// TIA Portal V17 export
// export: Created 2025-08-05T06:59:04.9381121Z, ExportSetting WithDefaults, DisplayName Totally Integrated Automation Portal, DisplayVersion V17 Update 5, DisplayName TIA Portal Openness, DisplayVersion V17 Update 5, DisplayName TIA Portal Version Control Interface, DisplayVersion V17, DisplayName SINAMICS Startdrive Advanced, DisplayVersion V17, DisplayName SINAMICS Startdrive G130, G150, S120, S150, SINAMICS MV, S210, DisplayVersion V17, DisplayName SINAMICS Startdrive G110M, G120, G120C, G120D, G120P, G115D, DisplayVersion V17, DisplayName STEP 7 Professional, DisplayVersion V17 Update 5, DisplayName STEP 7 Safety, DisplayVersion V17, DisplayName WinCC Advanced, DisplayVersion V17 Update 5
FUNCTION_BLOCK "FB_CentreStand_Fix_Seq_7"   // FB1, LAD
VERSION : 0.1
// stored: AutoNumber true, IsIECCheckEnabled false, UDAEnableTagReadback false
   VAR_INPUT
      iAutoRunning : Bool;
      iFixClamp : Bool;
      iFixEmpty : Bool;
      iFixTrayPresent : Bool;
      iFixUnclamp : Bool;
      iR1DropOver : Bool;
      iR1PickOver : Bool;
      iR2OperationOver : Bool;
      iR2ServiceActivated : Bool;
      iR2ServiceCompleted : Bool;
      iReset_fault : Bool;
      iRobotOutofZone : Bool;
      iSstMode : Bool;
      iSstPB : Bool;
   END_VAR
   VAR_OUTPUT
      qFixClamp : Bool;
      qFixUnclamp : Bool;
      qR1ReadytoDropTray : Bool;
      qR1ReadytoPickTray : Bool;
      qR2OperationStart : Bool;
   END_VAR
   VAR_IN_OUT
      iqR2ServiceActive : Bool;
      iqR2ServiceCompleted : Bool;
   END_VAR
   VAR DB_SPECIFIC
      StateNo : Int;
      s138_WaitBothRbtOutAl : Bool;
      s138_WaitBothRbtOutAl_T1 : Bool;
      s138_WaitBothRbtOutAl_T2 : Bool;
      s139_FixEmpty : Bool;
      s139_FixEmpty_T1 : Bool;
      s140_FixTrayPrsntRec : Bool;
      s140_FixTrayPrsntRec_T1 : Bool;
      s140_FixTrayPrsntRec_T2 : Bool;
      s141_FixUnclampCmd : Bool;
      s141_FixUnclampCmd_T1 : Bool;
      s142_TrayRdyDropFix : Bool;
      s142_TrayRdyDropFix_T1 : Bool;
      s143_RbtDropFixChkTr : Bool;
      s143_RbtDropFixChkTr_T1 : Bool;
      s144_RbtOutAreaDrop : Bool;
      s144_RbtOutAreaDrop_T1 : Bool;
      s145_FixClamp : Bool;
      s145_FixClamp_T1 : Bool;
      s146_Rbt2AlloyOpOver : Bool;
      s146_Rbt2AlloyOpOver_T1 : Bool;
      s147_FixUnclmpCmdOvr : Bool;
      s147_FixUnclmpCmdOvr_T1 : Bool;
      s148_RdyPickTrayWait : Bool;
      s148_RdyPickTrayWait_T1 : Bool;
      s149_RbtPickTrayChkEm : Bool;
      s149_RbtPickTrayChkEm_T1 : Bool;
      s191_WaitRbt2OutArea : Bool;
      s191_WaitRbt2OutArea_T1 : Bool;
      sSst : Bool;
      sSstPulse : Bool;
      sSstRise : Bool;
      sStWtResetRel : Bool;
      sStWtResetRel_T1 : Bool;
   END_VAR
   VAR_TEMP
      tOne : Bool;
   END_VAR
   VAR_TEMP   // added for the SCL form of the ladder/FBD networks
      _w1 : Bool;
   END_VAR
BEGIN

REGION Network 1
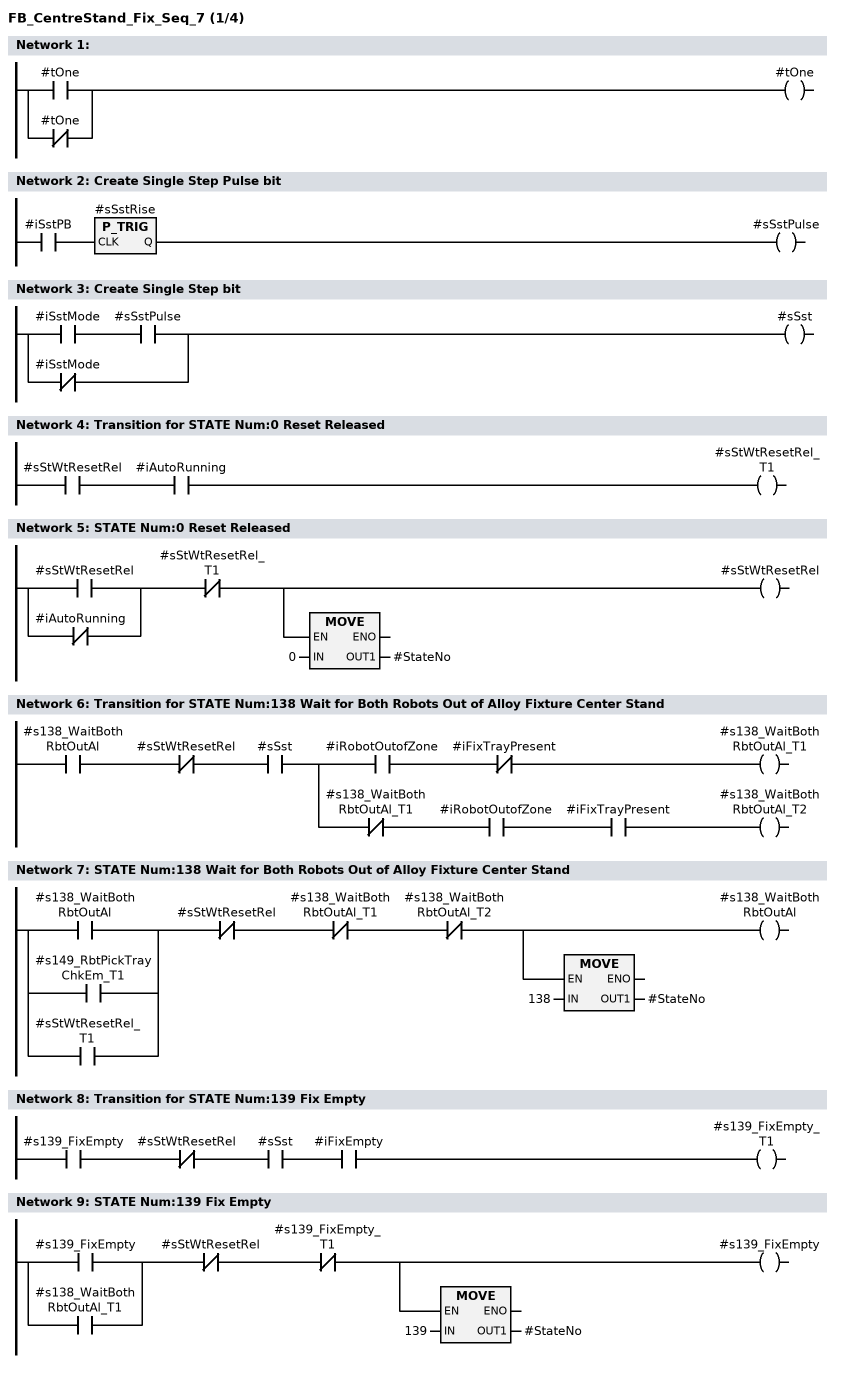
   RUNG wire#powerrail
      Contact( #tOne )
      wire#w1
      Coil( #tOne )
   END_RUNG
   RUNG wire#powerrail
      I_Contact( #tOne )
   END_RUNG wire#w1
   // the same network as SCL:
   #tOne := #tOne OR NOT #tOne;
END_REGION

REGION Network 2: Create Single Step Pulse bit
   RUNG wire#powerrail
      Contact( #iSstPB )
      P_Trig( #sSstRise )
      Coil( #sSstPulse )
   END_RUNG
   // the same network as SCL:
   #_w1 := #iSstPB AND NOT #sSstRise;   // rising edge
   #sSstRise := #iSstPB;
   #sSstPulse := #_w1;
END_REGION

REGION Network 3: Create Single Step bit
   RUNG wire#powerrail
      Contact( #iSstMode )
      Contact( #sSstPulse )
      wire#w1
      Coil( #sSst )
   END_RUNG
   RUNG wire#powerrail
      I_Contact( #iSstMode )
   END_RUNG wire#w1
   // the same network as SCL:
   #sSst := (#iSstMode AND #sSstPulse) OR NOT #iSstMode;
END_REGION

REGION Network 4: Transition for STATE Num:0 Reset Released
   RUNG wire#powerrail
      Contact( #sStWtResetRel )
      Contact( #iAutoRunning )
      Coil( #sStWtResetRel_T1 )
   END_RUNG
   // the same network as SCL:
   #sStWtResetRel_T1 := #sStWtResetRel AND #iAutoRunning;
END_REGION

REGION Network 5: STATE Num:0 Reset Released
   RUNG wire#powerrail
      Contact( #sStWtResetRel )
      wire#w1
      I_Contact( #sStWtResetRel_T1 )
      wire#w2
      Coil( #sStWtResetRel )
   END_RUNG
   RUNG wire#powerrail
      I_Contact( #iAutoRunning )
   END_RUNG wire#w1
   RUNG wire#w2
      { S7_GenerateENO := "TRUE" } Move(in := 0, out1 => #StateNo)
   END_RUNG
   // the same network as SCL:
   #sStWtResetRel := (#sStWtResetRel OR NOT #iAutoRunning) AND NOT #sStWtResetRel_T1;
   IF #sStWtResetRel THEN #StateNo := 0; END_IF;
END_REGION

REGION Network 6: Transition for STATE Num:138 Wait for Both Robots Out of Alloy Fixture Center Stand
   RUNG wire#powerrail
      Contact( #s138_WaitBothRbtOutAl )
      I_Contact( #sStWtResetRel )
      Contact( #sSst )
      wire#w1
      Contact( #iRobotOutofZone )
      I_Contact( #iFixTrayPresent )
      Coil( #s138_WaitBothRbtOutAl_T1 )
   END_RUNG
   RUNG wire#w1
      I_Contact( #s138_WaitBothRbtOutAl_T1 )
      Contact( #iRobotOutofZone )
      Contact( #iFixTrayPresent )
      Coil( #s138_WaitBothRbtOutAl_T2 )
   END_RUNG
   // the same network as SCL:
   #_w1 := #s138_WaitBothRbtOutAl AND NOT #sStWtResetRel AND #sSst;
   #s138_WaitBothRbtOutAl_T1 := #_w1 AND #iRobotOutofZone AND NOT #iFixTrayPresent;
   #s138_WaitBothRbtOutAl_T2 := #_w1 AND NOT #s138_WaitBothRbtOutAl_T1 AND #iRobotOutofZone AND #iFixTrayPresent;
END_REGION

REGION Network 7: STATE Num:138 Wait for Both Robots Out of Alloy Fixture Center Stand
   RUNG wire#powerrail
      Contact( #s138_WaitBothRbtOutAl )
      wire#w1
      I_Contact( #sStWtResetRel )
      I_Contact( #s138_WaitBothRbtOutAl_T1 )
      I_Contact( #s138_WaitBothRbtOutAl_T2 )
      wire#w2
      Coil( #s138_WaitBothRbtOutAl )
   END_RUNG
   RUNG wire#powerrail
      Contact( #s149_RbtPickTrayChkEm_T1 )
   END_RUNG wire#w1
   RUNG wire#powerrail
      Contact( #sStWtResetRel_T1 )
   END_RUNG wire#w1
   RUNG wire#w2
      { S7_GenerateENO := "TRUE" } Move(in := 138, out1 => #StateNo)
   END_RUNG
   // the same network as SCL:
   #s138_WaitBothRbtOutAl := (#s138_WaitBothRbtOutAl OR #s149_RbtPickTrayChkEm_T1 OR #sStWtResetRel_T1) AND NOT #sStWtResetRel AND NOT #s138_WaitBothRbtOutAl_T1 AND NOT #s138_WaitBothRbtOutAl_T2;
   IF #s138_WaitBothRbtOutAl THEN #StateNo := 138; END_IF;
END_REGION

REGION Network 8: Transition for STATE Num:139 Fix Empty
   RUNG wire#powerrail
      Contact( #s139_FixEmpty )
      I_Contact( #sStWtResetRel )
      Contact( #sSst )
      Contact( #iFixEmpty )
      Coil( #s139_FixEmpty_T1 )
   END_RUNG
   // the same network as SCL:
   #s139_FixEmpty_T1 := #s139_FixEmpty AND NOT #sStWtResetRel AND #sSst AND #iFixEmpty;
END_REGION

REGION Network 9: STATE Num:139 Fix Empty
   RUNG wire#powerrail
      Contact( #s139_FixEmpty )
      wire#w1
      I_Contact( #sStWtResetRel )
      I_Contact( #s139_FixEmpty_T1 )
      wire#w2
      Coil( #s139_FixEmpty )
   END_RUNG
   RUNG wire#powerrail
      Contact( #s138_WaitBothRbtOutAl_T1 )
   END_RUNG wire#w1
   RUNG wire#w2
      { S7_GenerateENO := "TRUE" } Move(in := 139, out1 => #StateNo)
   END_RUNG
   // the same network as SCL:
   #s139_FixEmpty := (#s139_FixEmpty OR #s138_WaitBothRbtOutAl_T1) AND NOT #sStWtResetRel AND NOT #s139_FixEmpty_T1;
   IF #s139_FixEmpty THEN #StateNo := 139; END_IF;
END_REGION

REGION Network 10: Transition for STATE Num:140 Fix Tray Present_Rec Operation pending
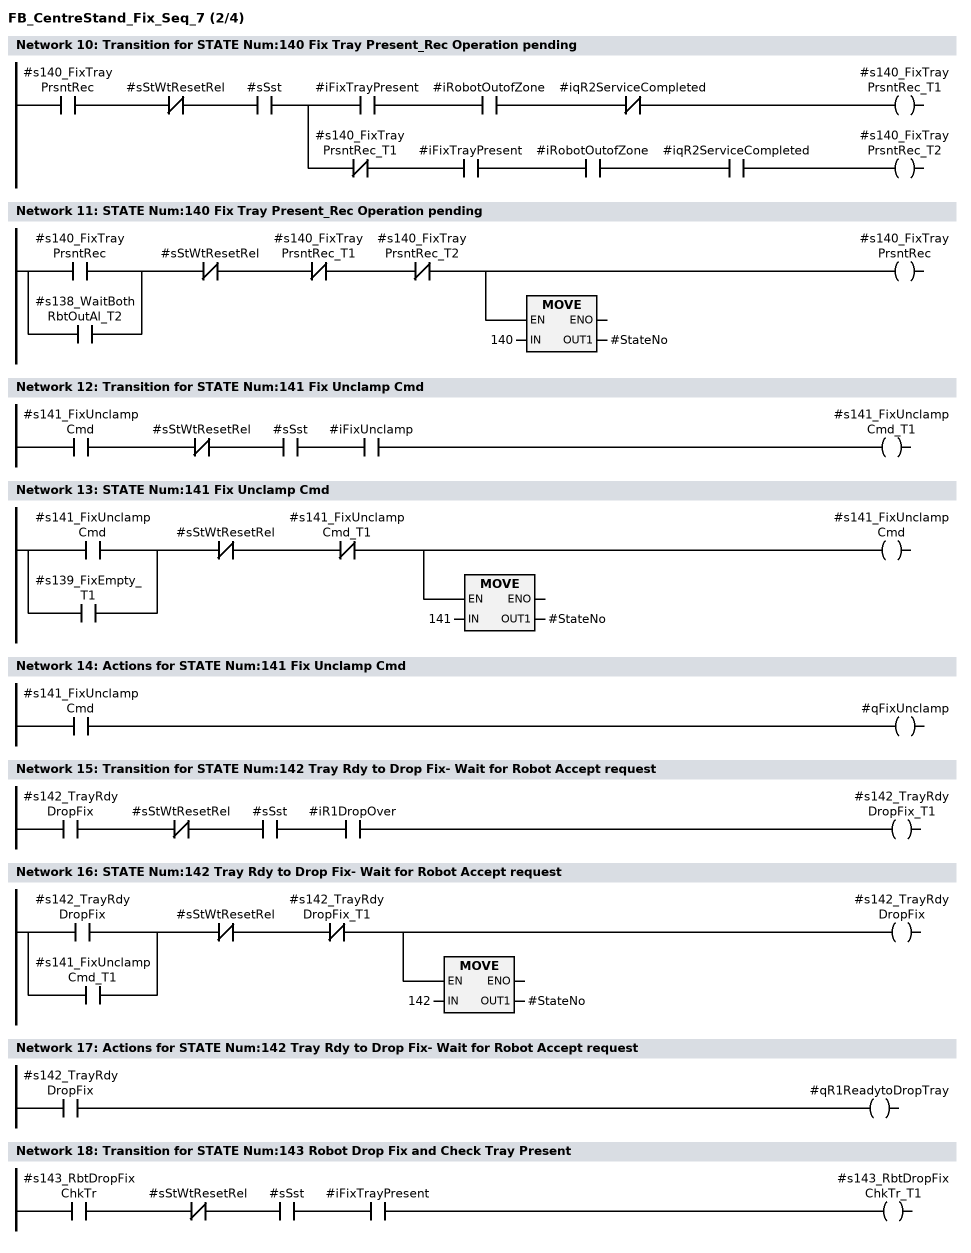
   RUNG wire#powerrail
      Contact( #s140_FixTrayPrsntRec )
      I_Contact( #sStWtResetRel )
      Contact( #sSst )
      wire#w1
      Contact( #iFixTrayPresent )
      Contact( #iRobotOutofZone )
      I_Contact( #iqR2ServiceCompleted )
      Coil( #s140_FixTrayPrsntRec_T1 )
   END_RUNG
   RUNG wire#w1
      I_Contact( #s140_FixTrayPrsntRec_T1 )
      Contact( #iFixTrayPresent )
      Contact( #iRobotOutofZone )
      Contact( #iqR2ServiceCompleted )
      Coil( #s140_FixTrayPrsntRec_T2 )
   END_RUNG
   // the same network as SCL:
   #_w1 := #s140_FixTrayPrsntRec AND NOT #sStWtResetRel AND #sSst;
   #s140_FixTrayPrsntRec_T1 := #_w1 AND #iFixTrayPresent AND #iRobotOutofZone AND NOT #iqR2ServiceCompleted;
   #s140_FixTrayPrsntRec_T2 := #_w1 AND NOT #s140_FixTrayPrsntRec_T1 AND #iFixTrayPresent AND #iRobotOutofZone AND #iqR2ServiceCompleted;
END_REGION

REGION Network 11: STATE Num:140 Fix Tray Present_Rec Operation pending
   RUNG wire#powerrail
      Contact( #s140_FixTrayPrsntRec )
      wire#w1
      I_Contact( #sStWtResetRel )
      I_Contact( #s140_FixTrayPrsntRec_T1 )
      I_Contact( #s140_FixTrayPrsntRec_T2 )
      wire#w2
      Coil( #s140_FixTrayPrsntRec )
   END_RUNG
   RUNG wire#powerrail
      Contact( #s138_WaitBothRbtOutAl_T2 )
   END_RUNG wire#w1
   RUNG wire#w2
      { S7_GenerateENO := "TRUE" } Move(in := 140, out1 => #StateNo)
   END_RUNG
   // the same network as SCL:
   #s140_FixTrayPrsntRec := (#s140_FixTrayPrsntRec OR #s138_WaitBothRbtOutAl_T2) AND NOT #sStWtResetRel AND NOT #s140_FixTrayPrsntRec_T1 AND NOT #s140_FixTrayPrsntRec_T2;
   IF #s140_FixTrayPrsntRec THEN #StateNo := 140; END_IF;
END_REGION

REGION Network 12: Transition for STATE Num:141 Fix Unclamp Cmd
   RUNG wire#powerrail
      Contact( #s141_FixUnclampCmd )
      I_Contact( #sStWtResetRel )
      Contact( #sSst )
      Contact( #iFixUnclamp )
      Coil( #s141_FixUnclampCmd_T1 )
   END_RUNG
   // the same network as SCL:
   #s141_FixUnclampCmd_T1 := #s141_FixUnclampCmd AND NOT #sStWtResetRel AND #sSst AND #iFixUnclamp;
END_REGION

REGION Network 13: STATE Num:141 Fix Unclamp Cmd
   RUNG wire#powerrail
      Contact( #s141_FixUnclampCmd )
      wire#w1
      I_Contact( #sStWtResetRel )
      I_Contact( #s141_FixUnclampCmd_T1 )
      wire#w2
      Coil( #s141_FixUnclampCmd )
   END_RUNG
   RUNG wire#powerrail
      Contact( #s139_FixEmpty_T1 )
   END_RUNG wire#w1
   RUNG wire#w2
      { S7_GenerateENO := "TRUE" } Move(in := 141, out1 => #StateNo)
   END_RUNG
   // the same network as SCL:
   #s141_FixUnclampCmd := (#s141_FixUnclampCmd OR #s139_FixEmpty_T1) AND NOT #sStWtResetRel AND NOT #s141_FixUnclampCmd_T1;
   IF #s141_FixUnclampCmd THEN #StateNo := 141; END_IF;
END_REGION

REGION Network 14: Actions for STATE Num:141 Fix Unclamp Cmd
   RUNG wire#powerrail
      Contact( #s141_FixUnclampCmd )
      Coil( #qFixUnclamp )
   END_RUNG
   // the same network as SCL:
   #qFixUnclamp := #s141_FixUnclampCmd;
END_REGION

REGION Network 15: Transition for STATE Num:142 Tray Rdy to Drop Fix- Wait for Robot Accept request
   RUNG wire#powerrail
      Contact( #s142_TrayRdyDropFix )
      I_Contact( #sStWtResetRel )
      Contact( #sSst )
      Contact( #iR1DropOver )
      Coil( #s142_TrayRdyDropFix_T1 )
   END_RUNG
   // the same network as SCL:
   #s142_TrayRdyDropFix_T1 := #s142_TrayRdyDropFix AND NOT #sStWtResetRel AND #sSst AND #iR1DropOver;
END_REGION

REGION Network 16: STATE Num:142 Tray Rdy to Drop Fix- Wait for Robot Accept request
   RUNG wire#powerrail
      Contact( #s142_TrayRdyDropFix )
      wire#w1
      I_Contact( #sStWtResetRel )
      I_Contact( #s142_TrayRdyDropFix_T1 )
      wire#w2
      Coil( #s142_TrayRdyDropFix )
   END_RUNG
   RUNG wire#powerrail
      Contact( #s141_FixUnclampCmd_T1 )
   END_RUNG wire#w1
   RUNG wire#w2
      { S7_GenerateENO := "TRUE" } Move(in := 142, out1 => #StateNo)
   END_RUNG
   // the same network as SCL:
   #s142_TrayRdyDropFix := (#s142_TrayRdyDropFix OR #s141_FixUnclampCmd_T1) AND NOT #sStWtResetRel AND NOT #s142_TrayRdyDropFix_T1;
   IF #s142_TrayRdyDropFix THEN #StateNo := 142; END_IF;
END_REGION

REGION Network 17: Actions for STATE Num:142 Tray Rdy to Drop Fix- Wait for Robot Accept request
   RUNG wire#powerrail
      Contact( #s142_TrayRdyDropFix )
      Coil( #qR1ReadytoDropTray )
   END_RUNG
   // the same network as SCL:
   #qR1ReadytoDropTray := #s142_TrayRdyDropFix;
END_REGION

REGION Network 18: Transition for STATE Num:143 Robot Drop Fix and Check Tray Present
   RUNG wire#powerrail
      Contact( #s143_RbtDropFixChkTr )
      I_Contact( #sStWtResetRel )
      Contact( #sSst )
      Contact( #iFixTrayPresent )
      Coil( #s143_RbtDropFixChkTr_T1 )
   END_RUNG
   // the same network as SCL:
   #s143_RbtDropFixChkTr_T1 := #s143_RbtDropFixChkTr AND NOT #sStWtResetRel AND #sSst AND #iFixTrayPresent;
END_REGION

REGION Network 19: STATE Num:143 Robot Drop Fix and Check Tray Present
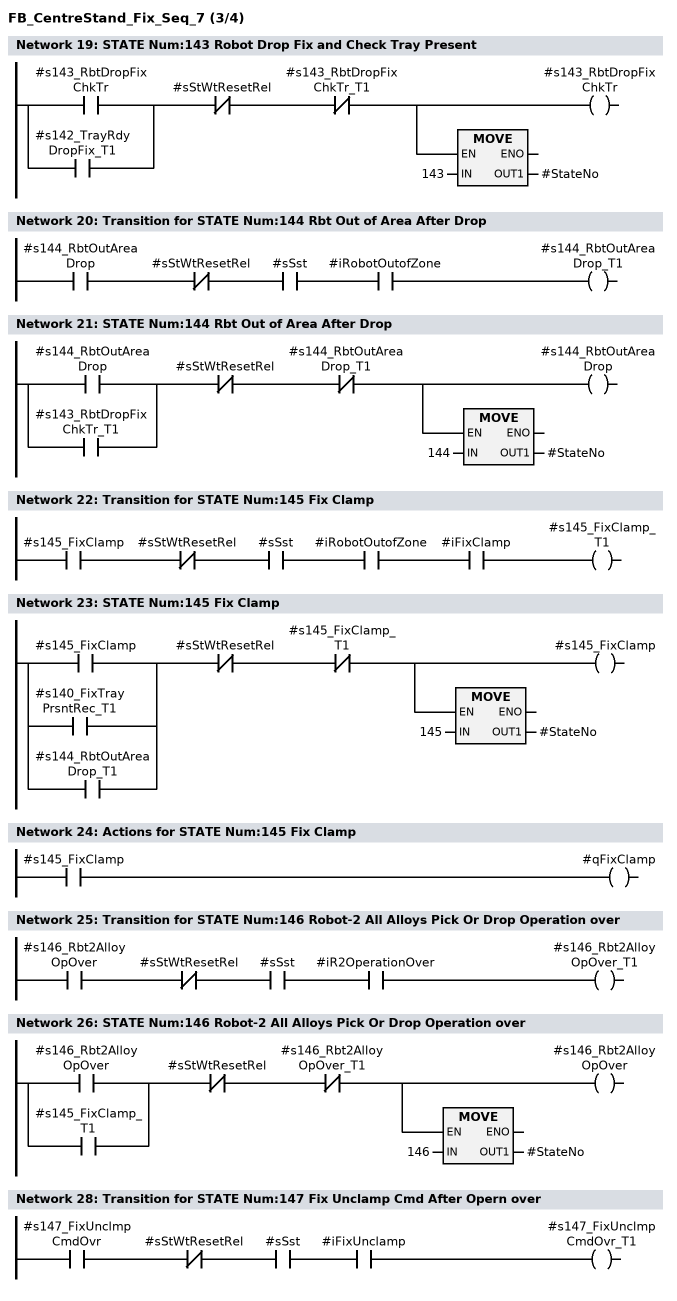
   RUNG wire#powerrail
      Contact( #s143_RbtDropFixChkTr )
      wire#w1
      I_Contact( #sStWtResetRel )
      I_Contact( #s143_RbtDropFixChkTr_T1 )
      wire#w2
      Coil( #s143_RbtDropFixChkTr )
   END_RUNG
   RUNG wire#powerrail
      Contact( #s142_TrayRdyDropFix_T1 )
   END_RUNG wire#w1
   RUNG wire#w2
      { S7_GenerateENO := "TRUE" } Move(in := 143, out1 => #StateNo)
   END_RUNG
   // the same network as SCL:
   #s143_RbtDropFixChkTr := (#s143_RbtDropFixChkTr OR #s142_TrayRdyDropFix_T1) AND NOT #sStWtResetRel AND NOT #s143_RbtDropFixChkTr_T1;
   IF #s143_RbtDropFixChkTr THEN #StateNo := 143; END_IF;
END_REGION

REGION Network 20: Transition for STATE Num:144 Rbt Out of Area After Drop
   RUNG wire#powerrail
      Contact( #s144_RbtOutAreaDrop )
      I_Contact( #sStWtResetRel )
      Contact( #sSst )
      Contact( #iRobotOutofZone )
      Coil( #s144_RbtOutAreaDrop_T1 )
   END_RUNG
   // the same network as SCL:
   #s144_RbtOutAreaDrop_T1 := #s144_RbtOutAreaDrop AND NOT #sStWtResetRel AND #sSst AND #iRobotOutofZone;
END_REGION

REGION Network 21: STATE Num:144 Rbt Out of Area After Drop
   RUNG wire#powerrail
      Contact( #s144_RbtOutAreaDrop )
      wire#w1
      I_Contact( #sStWtResetRel )
      I_Contact( #s144_RbtOutAreaDrop_T1 )
      wire#w2
      Coil( #s144_RbtOutAreaDrop )
   END_RUNG
   RUNG wire#powerrail
      Contact( #s143_RbtDropFixChkTr_T1 )
   END_RUNG wire#w1
   RUNG wire#w2
      { S7_GenerateENO := "TRUE" } Move(in := 144, out1 => #StateNo)
   END_RUNG
   // the same network as SCL:
   #s144_RbtOutAreaDrop := (#s144_RbtOutAreaDrop OR #s143_RbtDropFixChkTr_T1) AND NOT #sStWtResetRel AND NOT #s144_RbtOutAreaDrop_T1;
   IF #s144_RbtOutAreaDrop THEN #StateNo := 144; END_IF;
END_REGION

REGION Network 22: Transition for STATE Num:145 Fix Clamp
   RUNG wire#powerrail
      Contact( #s145_FixClamp )
      I_Contact( #sStWtResetRel )
      Contact( #sSst )
      Contact( #iRobotOutofZone )
      Contact( #iFixClamp )
      Coil( #s145_FixClamp_T1 )
   END_RUNG
   // the same network as SCL:
   #s145_FixClamp_T1 := #s145_FixClamp AND NOT #sStWtResetRel AND #sSst AND #iRobotOutofZone AND #iFixClamp;
END_REGION

REGION Network 23: STATE Num:145 Fix Clamp
   RUNG wire#powerrail
      Contact( #s145_FixClamp )
      wire#w1
      I_Contact( #sStWtResetRel )
      I_Contact( #s145_FixClamp_T1 )
      wire#w2
      Coil( #s145_FixClamp )
   END_RUNG
   RUNG wire#powerrail
      Contact( #s140_FixTrayPrsntRec_T1 )
   END_RUNG wire#w1
   RUNG wire#powerrail
      Contact( #s144_RbtOutAreaDrop_T1 )
   END_RUNG wire#w1
   RUNG wire#w2
      { S7_GenerateENO := "TRUE" } Move(in := 145, out1 => #StateNo)
   END_RUNG
   // the same network as SCL:
   #s145_FixClamp := (#s145_FixClamp OR #s140_FixTrayPrsntRec_T1 OR #s144_RbtOutAreaDrop_T1) AND NOT #sStWtResetRel AND NOT #s145_FixClamp_T1;
   IF #s145_FixClamp THEN #StateNo := 145; END_IF;
END_REGION

REGION Network 24: Actions for STATE Num:145 Fix Clamp
   RUNG wire#powerrail
      Contact( #s145_FixClamp )
      Coil( #qFixClamp )
   END_RUNG
   // the same network as SCL:
   #qFixClamp := #s145_FixClamp;
END_REGION

REGION Network 25: Transition for STATE Num:146 Robot-2 All Alloys Pick Or Drop Operation over
   RUNG wire#powerrail
      Contact( #s146_Rbt2AlloyOpOver )
      I_Contact( #sStWtResetRel )
      Contact( #sSst )
      Contact( #iR2OperationOver )
      Coil( #s146_Rbt2AlloyOpOver_T1 )
   END_RUNG
   // the same network as SCL:
   #s146_Rbt2AlloyOpOver_T1 := #s146_Rbt2AlloyOpOver AND NOT #sStWtResetRel AND #sSst AND #iR2OperationOver;
END_REGION

REGION Network 26: STATE Num:146 Robot-2 All Alloys Pick Or Drop Operation over
   RUNG wire#powerrail
      Contact( #s146_Rbt2AlloyOpOver )
      wire#w1
      I_Contact( #sStWtResetRel )
      I_Contact( #s146_Rbt2AlloyOpOver_T1 )
      wire#w2
      Coil( #s146_Rbt2AlloyOpOver )
   END_RUNG
   RUNG wire#powerrail
      Contact( #s145_FixClamp_T1 )
   END_RUNG wire#w1
   RUNG wire#w2
      { S7_GenerateENO := "TRUE" } Move(in := 146, out1 => #StateNo)
   END_RUNG
   // the same network as SCL:
   #s146_Rbt2AlloyOpOver := (#s146_Rbt2AlloyOpOver OR #s145_FixClamp_T1) AND NOT #sStWtResetRel AND NOT #s146_Rbt2AlloyOpOver_T1;
   IF #s146_Rbt2AlloyOpOver THEN #StateNo := 146; END_IF;
END_REGION

NETWORK
TITLE = Actions for STATE Num:146 Robot-2 All Alloys Pick Or Drop Operation over
      A     #s146_Rbt2AlloyOpOver;
      =     #qR2OperationStart;
      A     #iR2ServiceActivated;
      S     #iqR2ServiceActive;
      A     #iR2OperationOver;
      A     #iqR2ServiceActive;
      R     #iqR2ServiceActive;

REGION Network 28: Transition for STATE Num:147 Fix Unclamp Cmd After Opern over
   RUNG wire#powerrail
      Contact( #s147_FixUnclmpCmdOvr )
      I_Contact( #sStWtResetRel )
      Contact( #sSst )
      Contact( #iFixUnclamp )
      Coil( #s147_FixUnclmpCmdOvr_T1 )
   END_RUNG
   // the same network as SCL:
   #s147_FixUnclmpCmdOvr_T1 := #s147_FixUnclmpCmdOvr AND NOT #sStWtResetRel AND #sSst AND #iFixUnclamp;
END_REGION

REGION Network 29: STATE Num:147 Fix Unclamp Cmd After Opern over
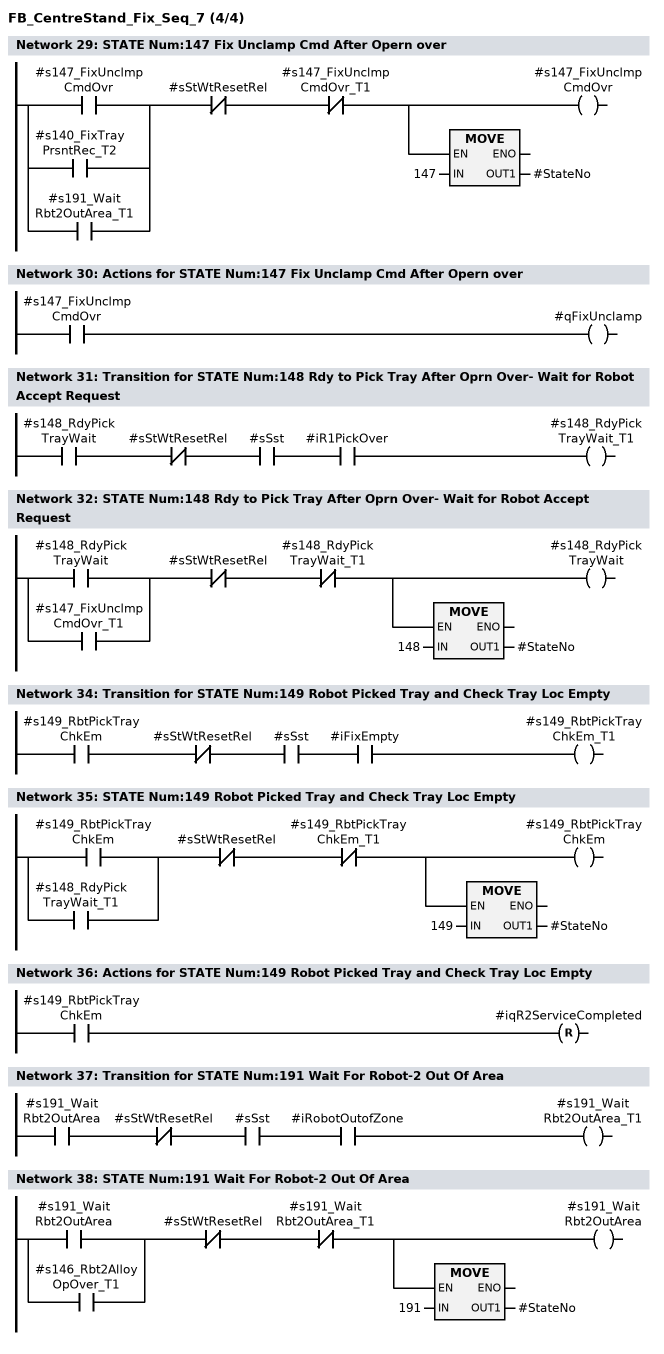
   RUNG wire#powerrail
      Contact( #s147_FixUnclmpCmdOvr )
      wire#w1
      I_Contact( #sStWtResetRel )
      I_Contact( #s147_FixUnclmpCmdOvr_T1 )
      wire#w2
      Coil( #s147_FixUnclmpCmdOvr )
   END_RUNG
   RUNG wire#powerrail
      Contact( #s140_FixTrayPrsntRec_T2 )
   END_RUNG wire#w1
   RUNG wire#powerrail
      Contact( #s191_WaitRbt2OutArea_T1 )
   END_RUNG wire#w1
   RUNG wire#w2
      { S7_GenerateENO := "TRUE" } Move(in := 147, out1 => #StateNo)
   END_RUNG
   // the same network as SCL:
   #s147_FixUnclmpCmdOvr := (#s147_FixUnclmpCmdOvr OR #s140_FixTrayPrsntRec_T2 OR #s191_WaitRbt2OutArea_T1) AND NOT #sStWtResetRel AND NOT #s147_FixUnclmpCmdOvr_T1;
   IF #s147_FixUnclmpCmdOvr THEN #StateNo := 147; END_IF;
END_REGION

REGION Network 30: Actions for STATE Num:147 Fix Unclamp Cmd After Opern over
   RUNG wire#powerrail
      Contact( #s147_FixUnclmpCmdOvr )
      Coil( #qFixUnclamp )
   END_RUNG
   // the same network as SCL:
   #qFixUnclamp := #s147_FixUnclmpCmdOvr;
END_REGION

REGION Network 31: Transition for STATE Num:148 Rdy to Pick Tray After Oprn Over- Wait for Robot Accept Request
   RUNG wire#powerrail
      Contact( #s148_RdyPickTrayWait )
      I_Contact( #sStWtResetRel )
      Contact( #sSst )
      Contact( #iR1PickOver )
      Coil( #s148_RdyPickTrayWait_T1 )
   END_RUNG
   // the same network as SCL:
   #s148_RdyPickTrayWait_T1 := #s148_RdyPickTrayWait AND NOT #sStWtResetRel AND #sSst AND #iR1PickOver;
END_REGION

REGION Network 32: STATE Num:148 Rdy to Pick Tray After Oprn Over- Wait for Robot Accept Request
   RUNG wire#powerrail
      Contact( #s148_RdyPickTrayWait )
      wire#w1
      I_Contact( #sStWtResetRel )
      I_Contact( #s148_RdyPickTrayWait_T1 )
      wire#w2
      Coil( #s148_RdyPickTrayWait )
   END_RUNG
   RUNG wire#powerrail
      Contact( #s147_FixUnclmpCmdOvr_T1 )
   END_RUNG wire#w1
   RUNG wire#w2
      { S7_GenerateENO := "TRUE" } Move(in := 148, out1 => #StateNo)
   END_RUNG
   // the same network as SCL:
   #s148_RdyPickTrayWait := (#s148_RdyPickTrayWait OR #s147_FixUnclmpCmdOvr_T1) AND NOT #sStWtResetRel AND NOT #s148_RdyPickTrayWait_T1;
   IF #s148_RdyPickTrayWait THEN #StateNo := 148; END_IF;
END_REGION

NETWORK
TITLE = Actions for STATE Num:148 Rdy to Pick Tray After Oprn Over- Wait for Robot Accept Request
      A     #s148_RdyPickTrayWait;
      =     #qR1ReadytoPickTray;
      A     #iR1PickOver;
      R     #iqR2ServiceCompleted;

REGION Network 34: Transition for STATE Num:149 Robot Picked Tray and Check Tray Loc Empty
   RUNG wire#powerrail
      Contact( #s149_RbtPickTrayChkEm )
      I_Contact( #sStWtResetRel )
      Contact( #sSst )
      Contact( #iFixEmpty )
      Coil( #s149_RbtPickTrayChkEm_T1 )
   END_RUNG
   // the same network as SCL:
   #s149_RbtPickTrayChkEm_T1 := #s149_RbtPickTrayChkEm AND NOT #sStWtResetRel AND #sSst AND #iFixEmpty;
END_REGION

REGION Network 35: STATE Num:149 Robot Picked Tray and Check Tray Loc Empty
   RUNG wire#powerrail
      Contact( #s149_RbtPickTrayChkEm )
      wire#w1
      I_Contact( #sStWtResetRel )
      I_Contact( #s149_RbtPickTrayChkEm_T1 )
      wire#w2
      Coil( #s149_RbtPickTrayChkEm )
   END_RUNG
   RUNG wire#powerrail
      Contact( #s148_RdyPickTrayWait_T1 )
   END_RUNG wire#w1
   RUNG wire#w2
      { S7_GenerateENO := "TRUE" } Move(in := 149, out1 => #StateNo)
   END_RUNG
   // the same network as SCL:
   #s149_RbtPickTrayChkEm := (#s149_RbtPickTrayChkEm OR #s148_RdyPickTrayWait_T1) AND NOT #sStWtResetRel AND NOT #s149_RbtPickTrayChkEm_T1;
   IF #s149_RbtPickTrayChkEm THEN #StateNo := 149; END_IF;
END_REGION

REGION Network 36: Actions for STATE Num:149 Robot Picked Tray and Check Tray Loc Empty
   RUNG wire#powerrail
      Contact( #s149_RbtPickTrayChkEm )
      R_Coil( #iqR2ServiceCompleted )
   END_RUNG
   // the same network as SCL:
   IF #s149_RbtPickTrayChkEm THEN #iqR2ServiceCompleted := FALSE; END_IF;
END_REGION

REGION Network 37: Transition for STATE Num:191 Wait For Robot-2 Out Of Area
   RUNG wire#powerrail
      Contact( #s191_WaitRbt2OutArea )
      I_Contact( #sStWtResetRel )
      Contact( #sSst )
      Contact( #iRobotOutofZone )
      Coil( #s191_WaitRbt2OutArea_T1 )
   END_RUNG
   // the same network as SCL:
   #s191_WaitRbt2OutArea_T1 := #s191_WaitRbt2OutArea AND NOT #sStWtResetRel AND #sSst AND #iRobotOutofZone;
END_REGION

REGION Network 38: STATE Num:191 Wait For Robot-2 Out Of Area
   RUNG wire#powerrail
      Contact( #s191_WaitRbt2OutArea )
      wire#w1
      I_Contact( #sStWtResetRel )
      I_Contact( #s191_WaitRbt2OutArea_T1 )
      wire#w2
      Coil( #s191_WaitRbt2OutArea )
   END_RUNG
   RUNG wire#powerrail
      Contact( #s146_Rbt2AlloyOpOver_T1 )
   END_RUNG wire#w1
   RUNG wire#w2
      { S7_GenerateENO := "TRUE" } Move(in := 191, out1 => #StateNo)
   END_RUNG
   // the same network as SCL:
   #s191_WaitRbt2OutArea := (#s191_WaitRbt2OutArea OR #s146_Rbt2AlloyOpOver_T1) AND NOT #sStWtResetRel AND NOT #s191_WaitRbt2OutArea_T1;
   IF #s191_WaitRbt2OutArea THEN #StateNo := 191; END_IF;
END_REGION
END_FUNCTION_BLOCK
